StartTest(TestName := 'Test_ComErrorClearedByAcknowledge');
group_2(Run := TRUE, ErrAck := FALSE); // T_SafeGroup
conn_2(InjectComError := FALSE, StartupTime := T#0S); // T_SafeConnection
group_2(Run := TRUE, ErrAck := FALSE); // T_SafeGroup
conn_2(InjectComError := FALSE, StartupTime := T#0S); // T_SafeConnection
group_2(Run := TRUE, ErrAck := FALSE); // T_SafeGroup
conn_2(InjectComError := FALSE, StartupTime := T#0S); // T_SafeConnection
group_2(Run := TRUE, ErrAck := FALSE); // T_SafeGroup
conn_2(InjectComError := FALSE, StartupTime := T#0S); // T_SafeConnection
group_2(Run := TRUE, ErrAck := FALSE); // T_SafeGroup
conn_2(InjectComError := FALSE, StartupTime := T#0S); // T_SafeConnection
group_2(Run := TRUE, ErrAck := FALSE); // T_SafeGroup
conn_2(InjectComError := TRUE, StartupTime := T#0S); // T_SafeConnection
AssertEquals_BOOL(Expected := TRUE, Actual := conn_2.ComError, Message := 'com error');
AssertEquals_BOOL(Expected := FALSE, Actual := conn_2.InDataState, Message := 'dropped out of Data');
AssertEquals_BYTE(Expected := BYTE#16#15, Actual := conn_2.Diag, Message := 'diag: watchdog code with the error bit');
group_2(Run := TRUE, ErrAck := FALSE); // T_SafeGroup
conn_2(InjectComError := FALSE, StartupTime := T#0S); // T_SafeConnection
AssertEquals_BYTE(Expected := TO_BYTE(E_SafeGroupState.Error), Actual := group_2.State, Message := 'group ERROR');
group_2(Run := TRUE, ErrAck := TRUE); // T_SafeGroup
conn_2(InjectComError := FALSE, StartupTime := T#0S); // T_SafeConnection
group_2(Run := TRUE, ErrAck := FALSE); // T_SafeGroup
conn_2(InjectComError := FALSE, StartupTime := T#0S); // T_SafeConnection
group_2(Run := TRUE, ErrAck := FALSE); // T_SafeGroup
conn_2(InjectComError := FALSE, StartupTime := T#0S); // T_SafeConnection
group_2(Run := TRUE, ErrAck := FALSE); // T_SafeGroup
conn_2(InjectComError := FALSE, StartupTime := T#0S); // T_SafeConnection
group_2(Run := TRUE, ErrAck := FALSE); // T_SafeGroup
conn_2(InjectComError := FALSE, StartupTime := T#0S); // T_SafeConnection
group_2(Run := TRUE, ErrAck := FALSE); // T_SafeGroup
conn_2(InjectComError := FALSE, StartupTime := T#0S); // T_SafeConnection
AssertEquals_BOOL(Expected := FALSE, Actual := conn_2.ComError, Message := 'error cleared');
AssertEquals_BOOL(Expected := TRUE, Actual := conn_2.InDataState, Message := 'restarted to Data');
FinishTest(TestName := 'Test_ComErrorClearedByAcknowledge');
END_METHOD

END_FUNCTION_BLOCK

// ---- Tests/T_SafeConnShutdown_Tests_CFC.TcPOU
    // CFC twin of T_SafeConnShutdown_Tests: the same tests drawn as CFC diagrams, the way a TwinSAFE project is authored.
    FUNCTION_BLOCK T_SafeConnShutdown_Tests_CFC EXTENDS T_SafeCfcTestSuite
    VAR
    // Test_DeactivateShutsDownConnection
    group_1 : T_SafeGroup;
    conn_1 : T_SafeConnection(group := group_1);
    fb_1 : T_SafeConnShutdown(group := group_1, connection := conn_1);
END_VAR

Test_DeactivateShutsDownConnection();

METHOD PRIVATE Test_DeactivateShutsDownConnection
// note: this text did not pass the execution check against the stored diagram
StartTest(TestName := 'Test_DeactivateShutsDownConnection');
group_1(Run := TRUE, ErrAck := FALSE); // T_SafeGroup
conn_1(StartupTime := T#0S); // T_SafeConnection
fb_1(Deactivate1 := FALSE); // T_SafeConnShutdown
group_1(Run := TRUE, ErrAck := FALSE); // T_SafeGroup
conn_1(StartupTime := T#0S); // T_SafeConnection
fb_1(Deactivate1 := FALSE); // T_SafeConnShutdown
group_1(Run := TRUE, ErrAck := FALSE); // T_SafeGroup
conn_1(StartupTime := T#0S); // T_SafeConnection
fb_1(Deactivate1 := FALSE); // T_SafeConnShutdown
group_1(Run := TRUE, ErrAck := FALSE); // T_SafeGroup
conn_1(StartupTime := T#0S); // T_SafeConnection
fb_1(Deactivate1 := FALSE); // T_SafeConnShutdown
group_1(Run := TRUE, ErrAck := FALSE); // T_SafeGroup
conn_1(StartupTime := T#0S); // T_SafeConnection
fb_1(Deactivate1 := FALSE); // T_SafeConnShutdown
AssertEquals_BOOL(Expected := FALSE, Actual := fb_1.Deactivated, Message := 'connection up');
group_1(Run := TRUE, ErrAck := FALSE); // T_SafeGroup
fb_1(Deactivate1 := TRUE); // T_SafeConnShutdown
conn_1(StartupTime := T#0S); // T_SafeConnection
fb_1(Deactivate1 := TRUE); // T_SafeConnShutdown
AssertEquals_BOOL(Expected := TRUE, Actual := conn_1.IsShutdown, Message := 'connection shut down');
AssertEquals_BOOL(Expected := TRUE, Actual := fb_1.Deactivated, Message := 'Deactivated output on');
group_1(Run := TRUE, ErrAck := FALSE); // T_SafeGroup
fb_1(Deactivate1 := FALSE); // T_SafeConnShutdown
conn_1(StartupTime := T#0S); // T_SafeConnection
group_1(Run := TRUE, ErrAck := FALSE); // T_SafeGroup
fb_1(Deactivate1 := FALSE); // T_SafeConnShutdown
conn_1(StartupTime := T#0S); // T_SafeConnection
group_1(Run := TRUE, ErrAck := FALSE); // T_SafeGroup
fb_1(Deactivate1 := FALSE); // T_SafeConnShutdown
conn_1(StartupTime := T#0S); // T_SafeConnection
group_1(Run := TRUE, ErrAck := FALSE); // T_SafeGroup
fb_1(Deactivate1 := FALSE); // T_SafeConnShutdown
conn_1(StartupTime := T#0S); // T_SafeConnection
group_1(Run := TRUE, ErrAck := FALSE); // T_SafeGroup
fb_1(Deactivate1 := FALSE); // T_SafeConnShutdown
conn_1(StartupTime := T#0S); // T_SafeConnection
group_1(Run := TRUE, ErrAck := FALSE); // T_SafeGroup
fb_1(Deactivate1 := FALSE); // T_SafeConnShutdown
conn_1(StartupTime := T#0S); // T_SafeConnection
AssertEquals_BOOL(Expected := TRUE, Actual := conn_1.InDataState, Message := 'connection re-established');
AssertEquals_BOOL(Expected := FALSE, Actual := fb_1.Deactivated, Message := 'Deactivated output off');
FinishTest(TestName := 'Test_DeactivateShutsDownConnection');
END_METHOD

END_FUNCTION_BLOCK

// ---- Tests/T_SafeGroup_Tests_CFC.TcPOU
    // CFC twin of T_SafeGroup_Tests: the same tests drawn as CFC diagrams, the way a TwinSAFE project is authored.
    FUNCTION_BLOCK T_SafeGroup_Tests_CFC EXTENDS T_SafeCfcTestSuite
    VAR
    // Test_StopWhenRunFalse
    group_1 : T_SafeGroup;
    fb_1 : T_SafeAnd(group := group_1);
    // Test_RunsFunctionBlocksWithoutConnections
    group_2 : T_SafeGroup;
    fb_2 : T_SafeAnd(group := group_2);
    // Test_FbErrorStopsGroupAndErrAckRecovers
    group_3 : T_SafeGroup;
    eStop_3 : T_SafeEStop(group := group_3);
    andFb_3 : T_SafeAnd(group := group_3);
    // Test_ConnectionStartupAndComError
    group_4 : T_SafeGroup;
    terminal_4 : T_SafeInputTerminal(group := group_4);
    t1a_4 : TON;
    t1b_4 : TON;
    t2b_4 : TON;
    trig1a_4 : R_TRIG;
    trig1b_4 : R_TRIG;
    trig2b_4 : R_TRIG;
    t3_4 : TON;
    trig3_4 : R_TRIG;
    t0_4 : TON;
    t1_4 : TON;
    t2_4 : TON;
    t4_4 : TON;
    trig0_4 : R_TRIG;
    trig1_4 : R_TRIG;
    trig2_4 : R_TRIG;
    trig4_4 : R_TRIG;
END_VAR

Test_StopWhenRunFalse();
Test_RunsFunctionBlocksWithoutConnections();
Test_FbErrorStopsGroupAndErrAckRecovers();
Test_ConnectionStartupAndComError();

METHOD PRIVATE Test_StopWhenRunFalse
// note: this text did not pass the execution check against the stored diagram
StartTest(TestName := 'Test_StopWhenRunFalse');
group_1(Run := FALSE, ErrAck := FALSE); // T_SafeGroup
fb_1(AndIn1 := TRUE, AndIn2 := TRUE); // T_SafeAnd
AssertEquals_BYTE(Expected := TO_BYTE(E_SafeGroupState.Stop), Actual := group_1.State, Message := 'group STOP');
AssertEquals_BYTE(Expected := TO_BYTE(E_SafeFbState.Stop), Actual := fb_1.State, Message := 'FB STOP');
AssertEquals_BOOL(Expected := FALSE, Actual := group_1.InRun, Message := 'InRun off');
FinishTest(TestName := 'Test_StopWhenRunFalse');
END_METHOD

METHOD PRIVATE Test_RunsFunctionBlocksWithoutConnections
// note: this text did not pass the execution check against the stored diagram
StartTest(TestName := 'Test_RunsFunctionBlocksWithoutConnections');
group_2(Run := TRUE, ErrAck := FALSE); // T_SafeGroup
fb_2(AndIn1 := TRUE, AndIn2 := TRUE); // T_SafeAnd
group_2(Run := TRUE, ErrAck := FALSE); // T_SafeGroup
fb_2(AndIn1 := TRUE, AndIn2 := TRUE); // T_SafeAnd
AssertEquals_BYTE(Expected := TO_BYTE(E_SafeGroupState.Run), Actual := group_2.State, Message := 'group RUN');
AssertEquals_BOOL(Expected := TRUE, Actual := fb_2.AndOut, Message := 'FB executed');
AssertEquals_BOOL(Expected := TRUE, Actual := group_2.FbRun, Message := 'all FBs running');
FinishTest(TestName := 'Test_RunsFunctionBlocksWithoutConnections');
END_METHOD

METHOD PRIVATE Test_FbErrorStopsGroupAndErrAckRecovers
// note: this text did not pass the execution check against the stored diagram
StartTest(TestName := 'Test_FbErrorStopsGroupAndErrAckRecovers');
group_3(Run := TRUE, ErrAck := FALSE); // T_SafeGroup
eStop_3(Restart := FALSE, EDM1 := FALSE, EStopIn1 := TRUE); // T_SafeEStop
andFb_3(AndIn1 := TRUE, AndIn2 := TRUE); // T_SafeAnd
group_3(Run := TRUE, ErrAck := FALSE); // T_SafeGroup
eStop_3(Restart := FALSE, EDM1 := FALSE, EStopIn1 := TRUE); // T_SafeEStop
andFb_3(AndIn1 := TRUE, AndIn2 := TRUE); // T_SafeAnd
AssertEquals_BOOL(Expected := TRUE, Actual := andFb_3.AndOut, Message := 'AND running before the error');
group_3(Run := TRUE, ErrAck := FALSE); // T_SafeGroup
eStop_3(Restart := TRUE, EDM1 := FALSE, EStopIn1 := TRUE); // T_SafeEStop
andFb_3(AndIn1 := TRUE, AndIn2 := TRUE); // T_SafeAnd
group_3(Run := TRUE, ErrAck := FALSE); // T_SafeGroup
eStop_3(Restart := FALSE, EDM1 := FALSE, EStopIn1 := TRUE); // T_SafeEStop
andFb_3(AndIn1 := TRUE, AndIn2 := TRUE); // T_SafeAnd
AssertEquals_BOOL(Expected := TRUE, Actual := group_3.FbErr, Message := 'FbErr');
AssertEquals_BYTE(Expected := TO_BYTE(E_SafeGroupState.Error), Actual := group_3.State, Message := 'group ERROR');
AssertEquals_BYTE(Expected := TO_BYTE(E_SafeGroupDiag.FbError), Actual := group_3.Diag, Message := 'group diag FBERROR');
AssertEquals_BOOL(Expected := FALSE, Actual := andFb_3.AndOut, Message := 'other FB outputs forced safe');
AssertEquals_BYTE(Expected := TO_BYTE(E_SafeFbState.Stop), Actual := andFb_3.State, Message := 'other FB STOP');
group_3(Run := TRUE, ErrAck := TRUE); // T_SafeGroup
eStop_3(Restart := FALSE, EDM1 := FALSE, EStopIn1 := TRUE); // T_SafeEStop
andFb_3(AndIn1 := TRUE, AndIn2 := TRUE); // T_SafeAnd
group_3(Run := TRUE, ErrAck := TRUE); // T_SafeGroup
eStop_3(Restart := FALSE, EDM1 := FALSE, EStopIn1 := TRUE); // T_SafeEStop
andFb_3(AndIn1 := TRUE, AndIn2 := TRUE); // T_SafeAnd
AssertEquals_BYTE(Expected := TO_BYTE(E_SafeGroupState.Reset), Actual := group_3.State, Message := 'group RESET while ErrAck 1');
group_3(Run := TRUE, ErrAck := FALSE); // T_SafeGroup
eStop_3(Restart := FALSE, EDM1 := FALSE, EStopIn1 := TRUE); // T_SafeEStop
andFb_3(AndIn1 := TRUE, AndIn2 := TRUE); // T_SafeAnd
group_3(Run := TRUE, ErrAck := FALSE); // T_SafeGroup
eStop_3(Restart := FALSE, EDM1 := FALSE, EStopIn1 := TRUE); // T_SafeEStop
andFb_3(AndIn1 := TRUE, AndIn2 := TRUE); // T_SafeAnd
AssertEquals_BYTE(Expected := TO_BYTE(E_SafeGroupState.Run), Actual := group_3.State, Message := 'group RUN after ErrAck');
AssertEquals_BOOL(Expected := TRUE, Actual := andFb_3.AndOut, Message := 'AND running again');
AssertEquals_BYTE(Expected := TO_BYTE(E_SafeFbState.Safe), Actual := eStop_3.State, Message := 'ESTOP back in SAFE awaiting restart');
FinishTest(TestName := 'Test_FbErrorStopsGroupAndErrAckRecovers');
END_METHOD

METHOD PRIVATE Test_ConnectionStartupAndComError
// note: this text did not pass the execution check against the stored diagram
StartTest(TestName := 'Test_ConnectionStartupAndComError');
t0_4(IN := TRUE, PT := T#20MS); // TON
trig0_4(CLK := t0_4.Q); // R_TRIG
t1a_4(IN := TRUE, PT := T#380MS); // TON
t1_4(IN := TRUE, PT := T#400MS); // TON
t1b_4(IN := t1_4.Q, PT := T#30MS); // TON
t2_4(IN := t1_4.Q, PT := T#50MS); // TON
t2b_4(IN := t2_4.Q, PT := T#20MS); // TON
t3_4(IN := t2_4.Q, PT := T#50MS); // TON
t4_4(IN := t3_4.Q, PT := T#400MS); // TON
trig1a_4(CLK := t1a_4.Q); // R_TRIG
trig1b_4(CLK := t1b_4.Q); // R_TRIG
trig1_4(CLK := t1_4.Q); // R_TRIG
trig2_4(CLK := t2_4.Q); // R_TRIG
trig2b_4(CLK := t2b_4.Q); // R_TRIG
trig3_4(CLK := t3_4.Q); // R_TRIG
trig4_4(CLK := t4_4.Q); // R_TRIG
group_4(Run := TRUE, ErrAck := t2_4.Q AND NOT t3_4.Q); // T_SafeGroup
terminal_4(InjectComError := trig1_4.Q, StartupTime := T#150MS); // T_SafeInputTerminal
IF trig0_4.Q THEN AssertEquals_BYTE(Expected := TO_BYTE(E_SafeGroupState.Start), Actual := group_4.State, Message := 'group START while the connection starts up'); END_IF
IF trig0_4.Q THEN AssertEquals_BOOL(Expected := TRUE, Actual := group_4.ComStartup, Message := 'ComStartup'); END_IF
IF trig1a_4.Q THEN AssertEquals_BYTE(Expected := TO_BYTE(E_SafeGroupState.Run), Actual := group_4.State, Message := 'group RUN once the connection is in Data'); END_IF
IF trig1b_4.Q THEN AssertEquals_BOOL(Expected := TRUE, Actual := group_4.ComErr, Message := 'ComErr'); END_IF
IF trig1b_4.Q THEN AssertEquals_BYTE(Expected := TO_BYTE(E_SafeGroupState.Error), Actual := group_4.State, Message := 'group ERROR'); END_IF
IF trig2b_4.Q THEN AssertEquals_BYTE(Expected := TO_BYTE(E_SafeGroupState.Reset), Actual := group_4.State, Message := 'group RESET'); END_IF
IF trig3_4.Q THEN AssertEquals_BYTE(Expected := TO_BYTE(E_SafeGroupState.Start), Actual := group_4.State, Message := 'group START again after ack'); END_IF
IF trig4_4.Q THEN AssertEquals_BYTE(Expected := TO_BYTE(E_SafeGroupState.Run), Actual := group_4.State, Message := 'group RUN after reconnection'); END_IF
IF trig4_4.Q THEN FinishTest(TestName := 'Test_ConnectionStartupAndComError'); END_IF
END_METHOD

END_FUNCTION_BLOCK

// ---- Tests/User_FB_Tests/T_SafePulse_UserFB_Tests_CFC.TcPOU
    // CFC twin of T_SafePulse_UserFB_Tests: the same tests drawn as CFC diagrams, the way a TwinSAFE project is authored.
    FUNCTION_BLOCK T_SafePulse_UserFB_Tests_CFC EXTENDS T_SafeCfcTestSuite
    VAR
    // Test_PulseForDelayTimeWhileInputHeld
    group_1 : T_SafeGroup;
    fb_1 : T_SafePulse_UserFB(group := group_1) := (Parameters := (DelayTime := T#100MS));
    trigStart_1 : R_TRIG;
    t1_1 : TON;
    t2_1 : TON;
    trig1_1 : R_TRIG;
    trig2_1 : R_TRIG;
    // Test_PulseEndsWhenInputDrops
    group_2 : T_SafeGroup;
    fb_2 : T_SafePulse_UserFB(group := group_2) := (Parameters := (DelayTime := T#100MS));
    // Test_StoppedGivesNoOutput
    group_3 : T_SafeGroup;
    fb_3 : T_SafePulse_UserFB(group := group_3) := (Parameters := (DelayTime := T#100MS));
    // Test_InnerBlocksJoinTheGroup
    group_4 : T_SafeGroup;
    fb_4 : T_SafePulse_UserFB(group := group_4);
END_VAR

Test_PulseForDelayTimeWhileInputHeld();
Test_PulseEndsWhenInputDrops();
Test_StoppedGivesNoOutput();
Test_InnerBlocksJoinTheGroup();

METHOD PRIVATE Test_InnerBlocksJoinTheGroup
StartTest(TestName := 'Test_InnerBlocksJoinTheGroup');
AssertEquals_UINT(Expected := 3, Actual := group_4.FunctionBlockCount, Message := 'composite and its two inner blocks registered');
FinishTest(TestName := 'Test_InnerBlocksJoinTheGroup');
END_METHOD

METHOD PRIVATE Test_PulseEndsWhenInputDrops
// note: this text did not pass the execution check against the stored diagram
StartTest(TestName := 'Test_PulseEndsWhenInputDrops');
group_2(Run := TRUE, ErrAck := FALSE); // T_SafeGroup
fb_2(TonIn1 := TRUE); // T_SafePulse_UserFB
AssertEquals_BOOL(Expected := TRUE, Actual := fb_2.TonOut, Message := 'pulse on');
fb_2(TonIn1 := FALSE); // T_SafePulse_UserFB
AssertEquals_BOOL(Expected := FALSE, Actual := fb_2.TonOut, Message := 'pulse cut off when the input drops');
FinishTest(TestName := 'Test_PulseEndsWhenInputDrops');
END_METHOD

METHOD PRIVATE Test_PulseForDelayTimeWhileInputHeld
// note: this text did not pass the execution check against the stored diagram
StartTest(TestName := 'Test_PulseForDelayTimeWhileInputHeld');
trigStart_1(CLK := TRUE); // R_TRIG
t1_1(IN := TRUE, PT := T#50MS); // TON
trig1_1(CLK := t1_1.Q); // R_TRIG
t2_1(IN := TRUE, PT := T#250MS); // TON
trig2_1(CLK := t2_1.Q); // R_TRIG
group_1(Run := TRUE, ErrAck := FALSE); // T_SafeGroup
fb_1(TonIn1 := TRUE); // T_SafePulse_UserFB
IF trigStart_1.Q THEN AssertEquals_BOOL(Expected := TRUE, Actual := fb_1.TonOut, Message := 'pulse starts with the input'); END_IF
IF trig1_1.Q THEN AssertEquals_BOOL(Expected := TRUE, Actual := fb_1.TonOut, Message := 'pulse still on inside the delay time'); END_IF
IF trig2_1.Q THEN AssertEquals_BOOL(Expected := FALSE, Actual := fb_1.TonOut, Message := 'pulse ends after the delay time'); END_IF
IF trig2_1.Q THEN
    fb_1(TonIn1 := FALSE); // T_SafePulse_UserFB
END_IF
IF trig2_1.Q THEN AssertEquals_BOOL(Expected := FALSE, Actual := fb_1.TonOut, Message := 'no output with the input off'); END_IF
IF trig2_1.Q THEN
    fb_1(TonIn1 := TRUE); // T_SafePulse_UserFB
END_IF
IF trig2_1.Q THEN AssertEquals_BOOL(Expected := TRUE, Actual := fb_1.TonOut, Message := 'a new pulse starts on the next rising edge'); END_IF
IF trig2_1.Q THEN FinishTest(TestName := 'Test_PulseForDelayTimeWhileInputHeld'); END_IF
END_METHOD

METHOD PRIVATE Test_StoppedGivesNoOutput
// note: this text did not pass the execution check against the stored diagram
StartTest(TestName := 'Test_StoppedGivesNoOutput');
group_3(Run := FALSE, ErrAck := FALSE); // T_SafeGroup
fb_3(TonIn1 := TRUE); // T_SafePulse_UserFB
AssertEquals_BOOL(Expected := FALSE, Actual := fb_3.TonOut, Message := 'no output while the group is stopped');
FinishTest(TestName := 'Test_StoppedGivesNoOutput');
END_METHOD

END_FUNCTION_BLOCK

// ---- Tests/User_FB_Tests/T_SafeRTrig_UserFB_Tests_CFC.TcPOU
    // CFC twin of T_SafeRTrig_UserFB_Tests: the same tests drawn as CFC diagrams, the way a TwinSAFE project is authored.
    FUNCTION_BLOCK T_SafeRTrig_UserFB_Tests_CFC EXTENDS T_SafeCfcTestSuite
    VAR
    // Test_TriggerForOneCycleOnRisingEdge
    group_1 : T_SafeGroup;
    fb_1 : T_SafeRTrig_UserFB(group := group_1);
    // Test_StoppedGivesNoOutput
    group_2 : T_SafeGroup;
    fb_2 : T_SafeRTrig_UserFB(group := group_2);
    // Test_InnerBlocksJoinTheGroup
    group_3 : T_SafeGroup;
    fb_3 : T_SafeRTrig_UserFB(group := group_3);
END_VAR

Test_TriggerForOneCycleOnRisingEdge();
Test_StoppedGivesNoOutput();
Test_InnerBlocksJoinTheGroup();

METHOD PRIVATE Test_InnerBlocksJoinTheGroup
StartTest(TestName := 'Test_InnerBlocksJoinTheGroup');
AssertEquals_UINT(Expected := 3, Actual := group_3.FunctionBlockCount, Message := 'composite and its two inner blocks registered');
FinishTest(TestName := 'Test_InnerBlocksJoinTheGroup');
END_METHOD

METHOD PRIVATE Test_StoppedGivesNoOutput
// note: this text did not pass the execution check against the stored diagram
StartTest(TestName := 'Test_StoppedGivesNoOutput');
group_2(Run := FALSE, ErrAck := FALSE); // T_SafeGroup
fb_2(Signal := TRUE); // T_SafeRTrig_UserFB
AssertEquals_BOOL(Expected := FALSE, Actual := fb_2.Trigger, Message := 'no output while the group is stopped');
FinishTest(TestName := 'Test_StoppedGivesNoOutput');
END_METHOD

METHOD PRIVATE Test_TriggerForOneCycleOnRisingEdge
// note: this text did not pass the execution check against the stored diagram
